Fanuc KAREL source: kd00061.KL

-- PROVISIONAL review KL for V1013-1; original PC SHA256 afb10bec612ea3b927820b2776bdd265ae8158d9a8fa1fa859a7568de97d324d
-- Incomplete behavior may be omitted. Consult companion uncertainty JSON. Do not deploy.
PROGRAM KD00061
%NOLOCKGROUP
VAR
  I : INTEGER
  J : INTEGER
  B : BOOLEAN
  R : REAL
  S : STRING[80]
BEGIN
  -- UNRESOLVED_PC offsets 5-18; opcodes 9D,81,18,9D,1B,9D,12,9D,13,04
  -- UNRESOLVED_PC offsets 23-27; opcodes 7F
END KD00061
